// Tests for FB_SweepStop, switching the uncalibrated axes off after a stop in the calibration sweep (#113).
FUNCTION_BLOCK FB_SweepStop_Tests EXTENDS TcUnit.FB_TestSuite
VAR
END_VAR

Disables_Uncalibrated_Axes_After_Three_Settled_Scans();
Calibrated_Axis_Stays_Enabled();
Waits_While_Homing_Runs();
Not_Settled_Restarts_The_Count();
No_Disable_Without_Arm();
Disable_Is_A_One_Scan_Pulse();
Cancel_Drops_The_Request();
ArmAll_Disables_Calibrated_Axes_Too();
ArmAll_Is_Idempotent();
ArmAll_Waits_For_The_Focus();
Arm_Ignores_OtherBusy();
Arm_Does_Not_Narrow_A_Pending_ArmAll();
Cancel_Clears_All_Mode();

METHOD PRIVATE Disables_Uncalibrated_Axes_After_Three_Settled_Scans
VAR
	fbSw	: FB_SweepStop;
	i		: INT;
END_VAR
TEST('Disables_Uncalibrated_Axes_After_Three_Settled_Scans');
fbSw.Arm();
FOR i := 1 TO 2 DO
fbSw(bSettled := TRUE, bHaCalibrated := FALSE, bDecCalibrated := FALSE, bHaHoming := FALSE, bDecHoming := FALSE);
END_FOR
AssertEquals_BOOL(Expected := FALSE, Actual := fbSw.bDisableHa, Message := 'two scans: not yet');
fbSw(bSettled := TRUE, bHaCalibrated := FALSE, bDecCalibrated := FALSE, bHaHoming := FALSE, bDecHoming := FALSE);
AssertEquals_BOOL(Expected := TRUE, Actual := fbSw.bDisableHa, Message := 'HA off');
AssertEquals_BOOL(Expected := TRUE, Actual := fbSw.bDisableDec, Message := 'Dec off');
TEST_FINISHED();
END_METHOD

METHOD PRIVATE Calibrated_Axis_Stays_Enabled
VAR
	fbSw	: FB_SweepStop;
	i		: INT;
END_VAR
TEST('Calibrated_Axis_Stays_Enabled');
fbSw.Arm();
FOR i := 1 TO 3 DO
fbSw(bSettled := TRUE, bHaCalibrated := TRUE, bDecCalibrated := FALSE, bHaHoming := FALSE, bDecHoming := FALSE);
END_FOR
AssertEquals_BOOL(Expected := FALSE, Actual := fbSw.bDisableHa, Message := 'HA calibrated');
AssertEquals_BOOL(Expected := TRUE, Actual := fbSw.bDisableDec, Message := 'Dec off');
TEST_FINISHED();
END_METHOD

METHOD PRIVATE Waits_While_Homing_Runs
VAR
	fbSw	: FB_SweepStop;
	i		: INT;
END_VAR
TEST('Waits_While_Homing_Runs');
fbSw.Arm();
FOR i := 1 TO 50 DO
fbSw(bSettled := TRUE, bHaCalibrated := FALSE, bDecCalibrated := FALSE, bHaHoming := TRUE, bDecHoming := FALSE);
END_FOR
AssertEquals_BOOL(Expected := FALSE, Actual := fbSw.bDisableHa, Message := 'HA homing busy');
FOR i := 1 TO 50 DO
fbSw(bSettled := TRUE, bHaCalibrated := FALSE, bDecCalibrated := FALSE, bHaHoming := FALSE, bDecHoming := TRUE);
END_FOR
AssertEquals_BOOL(Expected := FALSE, Actual := fbSw.bDisableDec, Message := 'Dec homing busy');
FOR i := 1 TO 3 DO
fbSw(bSettled := TRUE, bHaCalibrated := FALSE, bDecCalibrated := FALSE, bHaHoming := FALSE, bDecHoming := FALSE);
END_FOR
AssertEquals_BOOL(Expected := TRUE, Actual := fbSw.bDisableHa, Message := 'off when the homing is idle');
TEST_FINISHED();
END_METHOD

METHOD PRIVATE Not_Settled_Restarts_The_Count
VAR
	fbSw	: FB_SweepStop;
	i		: INT;
END_VAR
TEST('Not_Settled_Restarts_The_Count');
fbSw.Arm();
FOR i := 1 TO 2 DO
fbSw(bSettled := TRUE, bHaCalibrated := FALSE, bDecCalibrated := FALSE, bHaHoming := FALSE, bDecHoming := FALSE);
END_FOR
fbSw(bSettled := FALSE, bHaCalibrated := FALSE, bDecCalibrated := FALSE, bHaHoming := FALSE, bDecHoming := FALSE);
FOR i := 1 TO 2 DO
fbSw(bSettled := TRUE, bHaCalibrated := FALSE, bDecCalibrated := FALSE, bHaHoming := FALSE, bDecHoming := FALSE);
END_FOR
AssertEquals_BOOL(Expected := FALSE, Actual := fbSw.bDisableHa, Message := 'count restarted');
fbSw(bSettled := TRUE, bHaCalibrated := FALSE, bDecCalibrated := FALSE, bHaHoming := FALSE, bDecHoming := FALSE);
AssertEquals_BOOL(Expected := TRUE, Actual := fbSw.bDisableHa, Message := 'off');
TEST_FINISHED();
END_METHOD

METHOD PRIVATE No_Disable_Without_Arm
VAR
	fbSw	: FB_SweepStop;
	i		: INT;
END_VAR
TEST('No_Disable_Without_Arm');
FOR i := 1 TO 20 DO
fbSw(bSettled := TRUE, bHaCalibrated := FALSE, bDecCalibrated := FALSE, bHaHoming := FALSE, bDecHoming := FALSE);
END_FOR
AssertEquals_BOOL(Expected := FALSE, Actual := fbSw.bDisableHa, Message := 'not armed');
AssertEquals_BOOL(Expected := FALSE, Actual := fbSw.bDisableDec, Message := 'not armed');
TEST_FINISHED();
END_METHOD

METHOD PRIVATE Disable_Is_A_One_Scan_Pulse
VAR
	fbSw	: FB_SweepStop;
	i		: INT;
END_VAR
TEST('Disable_Is_A_One_Scan_Pulse');
fbSw.Arm();
FOR i := 1 TO 3 DO
fbSw(bSettled := TRUE, bHaCalibrated := FALSE, bDecCalibrated := FALSE, bHaHoming := FALSE, bDecHoming := FALSE);
END_FOR
AssertEquals_BOOL(Expected := TRUE, Actual := fbSw.bDisableHa, Message := 'pulse');
fbSw(bSettled := TRUE, bHaCalibrated := FALSE, bDecCalibrated := FALSE, bHaHoming := FALSE, bDecHoming := FALSE);
AssertEquals_BOOL(Expected := FALSE, Actual := fbSw.bDisableHa, Message := 'only once');
AssertEquals_BOOL(Expected := FALSE, Actual := fbSw.bDisableDec, Message := 'only once');
TEST_FINISHED();
END_METHOD

METHOD PRIVATE Cancel_Drops_The_Request
VAR
	fbSw	: FB_SweepStop;
	i		: INT;
END_VAR
TEST('Cancel_Drops_The_Request');
fbSw.Arm();
FOR i := 1 TO 2 DO
fbSw(bSettled := TRUE, bHaCalibrated := FALSE, bDecCalibrated := FALSE, bHaHoming := FALSE, bDecHoming := FALSE);
END_FOR
fbSw.Cancel();
FOR i := 1 TO 10 DO
fbSw(bSettled := TRUE, bHaCalibrated := FALSE, bDecCalibrated := FALSE, bHaHoming := FALSE, bDecHoming := FALSE);
END_FOR
AssertEquals_BOOL(Expected := FALSE, Actual := fbSw.bDisableHa, Message := 'cancelled');
TEST_FINISHED();
END_METHOD

// #197: a park without a completed power-on switches every axis off, calibrated or not
METHOD PRIVATE ArmAll_Disables_Calibrated_Axes_Too
VAR
	fbSw	: FB_SweepStop;
	i		: INT;
END_VAR
TEST('ArmAll_Disables_Calibrated_Axes_Too');
fbSw.ArmAll();
FOR i := 1 TO 2 DO
fbSw(bSettled := TRUE, bHaCalibrated := TRUE, bDecCalibrated := TRUE, bHaHoming := FALSE, bDecHoming := FALSE);
END_FOR
AssertEquals_BOOL(Expected := FALSE, Actual := fbSw.bDisableHa, Message := 'two scans: not yet');
fbSw(bSettled := TRUE, bHaCalibrated := TRUE, bDecCalibrated := TRUE, bHaHoming := FALSE, bDecHoming := FALSE);
AssertEquals_BOOL(Expected := TRUE, Actual := fbSw.bDisableHa, Message := 'HA off although calibrated');
AssertEquals_BOOL(Expected := TRUE, Actual := fbSw.bDisableDec, Message := 'Dec off although calibrated');
fbSw(bSettled := TRUE, bHaCalibrated := TRUE, bDecCalibrated := TRUE, bHaHoming := FALSE, bDecHoming := FALSE);
AssertEquals_BOOL(Expected := FALSE, Actual := fbSw.bDisableHa, Message := 'one scan only');
TEST_FINISHED();
END_METHOD

// #197: the arbitration calls ArmAll every scan
METHOD PRIVATE ArmAll_Is_Idempotent
VAR
	fbSw	: FB_SweepStop;
	i		: INT;
END_VAR
TEST('ArmAll_Is_Idempotent');
FOR i := 1 TO 2 DO
fbSw.ArmAll();
fbSw(bSettled := TRUE, bHaCalibrated := TRUE, bDecCalibrated := TRUE, bHaHoming := FALSE, bDecHoming := FALSE);
END_FOR
fbSw.ArmAll();
fbSw(bSettled := TRUE, bHaCalibrated := TRUE, bDecCalibrated := TRUE, bHaHoming := FALSE, bDecHoming := FALSE);
AssertEquals_BOOL(Expected := TRUE, Actual := fbSw.bDisableHa, Message := 'ArmAll every scan does not restart the count');
TEST_FINISHED();
END_METHOD

// #197: the focus must not be moving when the axes are switched off (#56)
METHOD PRIVATE ArmAll_Waits_For_The_Focus
VAR
	fbSw	: FB_SweepStop;
	i		: INT;
END_VAR
TEST('ArmAll_Waits_For_The_Focus');
fbSw.ArmAll();
FOR i := 1 TO 20 DO
fbSw(bSettled := TRUE, bHaCalibrated := TRUE, bDecCalibrated := TRUE, bHaHoming := FALSE, bDecHoming := FALSE, bOtherBusy := TRUE);
END_FOR
AssertEquals_BOOL(Expected := FALSE, Actual := fbSw.bDisableHa, Message := 'the focus is moving');
FOR i := 1 TO 3 DO
fbSw(bSettled := TRUE, bHaCalibrated := TRUE, bDecCalibrated := TRUE, bHaHoming := FALSE, bDecHoming := FALSE, bOtherBusy := FALSE);
END_FOR
AssertEquals_BOOL(Expected := TRUE, Actual := fbSw.bDisableDec, Message := 'off when the focus is at rest');
TEST_FINISHED();
END_METHOD

// #113 mode unchanged
METHOD PRIVATE Arm_Ignores_OtherBusy
VAR
	fbSw	: FB_SweepStop;
	i		: INT;
END_VAR
TEST('Arm_Ignores_OtherBusy');
fbSw.Arm();
FOR i := 1 TO 3 DO
fbSw(bSettled := TRUE, bHaCalibrated := FALSE, bDecCalibrated := TRUE, bHaHoming := FALSE, bDecHoming := FALSE, bOtherBusy := TRUE);
END_FOR
AssertEquals_BOOL(Expected := TRUE, Actual := fbSw.bDisableHa, Message := 'the stop of #113 does not wait for the focus');
AssertEquals_BOOL(Expected := FALSE, Actual := fbSw.bDisableDec, Message := 'calibrated axis stays on');
TEST_FINISHED();
END_METHOD

// a stop after the park request must not undo the all-axes mode
METHOD PRIVATE Arm_Does_Not_Narrow_A_Pending_ArmAll
VAR
	fbSw	: FB_SweepStop;
	i		: INT;
END_VAR
TEST('Arm_Does_Not_Narrow_A_Pending_ArmAll');
fbSw.ArmAll();
fbSw.Arm();
FOR i := 1 TO 3 DO
fbSw(bSettled := TRUE, bHaCalibrated := TRUE, bDecCalibrated := TRUE, bHaHoming := FALSE, bDecHoming := FALSE);
END_FOR
AssertEquals_BOOL(Expected := TRUE, Actual := fbSw.bDisableHa, Message := 'still the all-axes mode');
TEST_FINISHED();
END_METHOD

// Cancel drops the all-axes mode
METHOD PRIVATE Cancel_Clears_All_Mode
VAR
	fbSw	: FB_SweepStop;
	i		: INT;
END_VAR
TEST('Cancel_Clears_All_Mode');
fbSw.ArmAll();
fbSw.Cancel();
fbSw.Arm();
FOR i := 1 TO 3 DO
fbSw(bSettled := TRUE, bHaCalibrated := TRUE, bDecCalibrated := FALSE, bHaHoming := FALSE, bDecHoming := FALSE);
END_FOR
AssertEquals_BOOL(Expected := FALSE, Actual := fbSw.bDisableHa, Message := 'calibrated axis stays on after Cancel');
AssertEquals_BOOL(Expected := TRUE, Actual := fbSw.bDisableDec, Message := 'uncalibrated axis off');
TEST_FINISHED();
END_METHOD

END_FUNCTION_BLOCK

(* stored: Version 1.1.0.1, ProductVersion 3.1.4024.15
   POU FB_SweepStop_Tests: Id {ae0811a0-07de-4121-bb40-416ce921270b}, SpecialFunc None
   Method Disables_Uncalibrated_Axes_After_Three_Settled_Scans: Id {45680a00-18a4-4788-9e68-873e3787f22d}
   Method Calibrated_Axis_Stays_Enabled: Id {de6d524c-a539-4e2c-a08d-c0b739f42296}
   Method Waits_While_Homing_Runs: Id {4341cace-590f-4d1a-9d38-90d5d93b63d7}
   Method Not_Settled_Restarts_The_Count: Id {16c76841-c3be-4715-a28a-cd0d9cfd6e71}
   Method No_Disable_Without_Arm: Id {99ce0184-c5eb-4ee8-b433-6fc478582d46}
   Method Disable_Is_A_One_Scan_Pulse: Id {238880f9-cf37-4d08-94aa-95129d981330}
   Method Cancel_Drops_The_Request: Id {852635e7-cb64-48be-8436-c0f348566caa}
   Method ArmAll_Disables_Calibrated_Axes_Too: Id {a1f0c3d2-5b6e-4a71-8c94-0d2e7f3a1b01}
   Method ArmAll_Is_Idempotent: Id {a1f0c3d2-5b6e-4a71-8c94-0d2e7f3a1b02}
   Method ArmAll_Waits_For_The_Focus: Id {a1f0c3d2-5b6e-4a71-8c94-0d2e7f3a1b03}
   Method Arm_Ignores_OtherBusy: Id {a1f0c3d2-5b6e-4a71-8c94-0d2e7f3a1b04}
   Method Arm_Does_Not_Narrow_A_Pending_ArmAll: Id {a1f0c3d2-5b6e-4a71-8c94-0d2e7f3a1b05}
   Method Cancel_Clears_All_Mode: Id {a1f0c3d2-5b6e-4a71-8c94-0d2e7f3a1b06} *)
